(* IEC 61131-3 sources: volt/packages/volt-lsp-iec/test-corpus/awa-palletizer/Device/Plc Logic/Application/Library Manager/(unresolved)/base interfaces, 4 files *)

(* ---- TYPECLASS.dut ---- *)
TYPE TYPECLASS :
(
	TYPE_BOOL := 0,
	TYPE_BIT := 1,
	TYPE_BYTE := 2,
	TYPE_WORD := 3,
	TYPE_DWORD := 4,
	TYPE_LWORD := 5,
	TYPE_SINT := 6,
	TYPE_INT := 7,
	TYPE_DINT := 8,
	TYPE_LINT := 9,
	TYPE_USINT := 10,
	TYPE_UINT := 11,
	TYPE_UDINT := 12,
	TYPE_ULINT := 13,
	TYPE_REAL := 14,
	TYPE_LREAL := 15,
	TYPE_STRING := 16,
	TYPE_WSTRING := 17,
	TYPE_TIME := 18,
	TYPE_DATE := 19,
	TYPE_DATEANDTIME := 20,
	TYPE_TIMEOFDAY := 21,
	TYPE_POINTER := 22,
	TYPE_REFERENCE := 23,
	TYPE_SUBRANGE := 24,
	TYPE_ENUM := 25,
	TYPE_ARRAY := 26,
	TYPE_PARAMS := 27,
	TYPE_USERDEF := 28,
	TYPE_NONE := 29,
	TYPE_ANY := 30,
	TYPE_ANYBIT := 31,
	TYPE_ANYDATE := 32,
	TYPE_ANYINT := 33,
	TYPE_ANYNUM := 34,
	TYPE_ANYREAL := 35,
	TYPE_LAZY := 36,
	TYPE_LTIME := 37,
	TYPE_BITCONST := 38,
	TYPE_UXINT := 39,
	TYPE_XWORD := 40,
	TYPE_XINT := 41,
	TYPE_XSRTING := 42,
	TYPE_VARLENARRAY := 43,
	TYPE_ANYSTRING := 44,
	TYPE_VECTOR := 45,
	TYPE_LDATE := 46,
	TYPE_LDATEANDTIME := 47,
	TYPE_LTIMEOFDAY := 48,
	TYPE_INTERFACE := 16#F000
);
END_TYPE

(* ---- COMPONENTIDS.gvl ---- *)
VAR_GLOBAL
	CMPID_IECCODE : DWORD := 16#1000;
	CMPID_CMPSTARTOEM : DWORD := 16#2000;
	CMPID_CMPENDOEM : DWORD := 16#3FFF;
END_VAR

(* ---- INTERFACEIDS.gvl ---- *)
VAR_GLOBAL
	ITFID_IBASE : DWORD := 16#0;
	ITFID_ICMPSTARTOEM : DWORD := 16#2000;
	ITFID_ICMPENDOEM : DWORD := 16#3FFF;
END_VAR

(* ---- IBASE.itf ---- *)
INTERFACE IBASE
END_INTERFACE

METHOD FB_EXIT : BOOL
VAR_INPUT
	BINCOPYCODE : BOOL;
END_VAR
END_METHOD

METHOD RELEASE : DINT
END_METHOD

METHOD FB_REINIT : BOOL
END_METHOD

METHOD ADDREF : DINT
END_METHOD

METHOD QUERYINTERFACE : POINTER TO POINTER TO BYTE
VAR_INPUT
	IID : DWORD;
	PRESULT : POINTER TO UDINT;
END_VAR
END_METHOD

METHOD FB_INIT : BOOL
VAR_INPUT
	BINITRETAINS : BOOL;
	BINCOPYCODE : BOOL;
END_VAR
END_METHOD
